FUNCTION_BLOCK PID_SINGLE_UPDATE_SEQUENCE (* One tuning attempt between samples; native validation pending *)
  (* Standard: 61499-2 *)
  (* Version 0.1, 2026-10-24, Guilherme *)
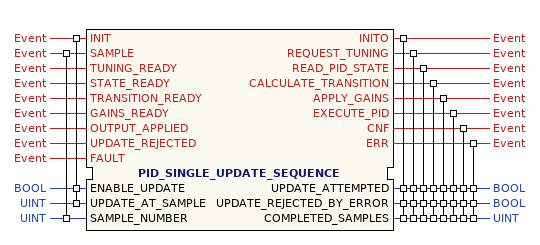
  EVENT_INPUT
    INIT WITH ENABLE_UPDATE, UPDATE_AT_SAMPLE;
    SAMPLE WITH SAMPLE_NUMBER;
    TUNING_READY;
    STATE_READY;
    TRANSITION_READY;
    GAINS_READY;
    OUTPUT_APPLIED;
    UPDATE_REJECTED;
    FAULT;
  END_EVENT
  EVENT_OUTPUT
    INITO WITH UPDATE_ATTEMPTED, UPDATE_REJECTED_BY_ERROR, COMPLETED_SAMPLES;
    REQUEST_TUNING WITH UPDATE_ATTEMPTED, UPDATE_REJECTED_BY_ERROR, COMPLETED_SAMPLES;
    READ_PID_STATE WITH UPDATE_ATTEMPTED, UPDATE_REJECTED_BY_ERROR, COMPLETED_SAMPLES;
    CALCULATE_TRANSITION WITH UPDATE_ATTEMPTED, UPDATE_REJECTED_BY_ERROR, COMPLETED_SAMPLES;
    APPLY_GAINS WITH UPDATE_ATTEMPTED, UPDATE_REJECTED_BY_ERROR, COMPLETED_SAMPLES;
    EXECUTE_PID WITH UPDATE_ATTEMPTED, UPDATE_REJECTED_BY_ERROR, COMPLETED_SAMPLES;
    CNF WITH UPDATE_ATTEMPTED, UPDATE_REJECTED_BY_ERROR, COMPLETED_SAMPLES;
    ERR WITH UPDATE_ATTEMPTED, UPDATE_REJECTED_BY_ERROR, COMPLETED_SAMPLES;
  END_EVENT
  VAR_INPUT
    ENABLE_UPDATE : BOOL;
    UPDATE_AT_SAMPLE : UINT;
    SAMPLE_NUMBER : UINT;
  END_VAR
  VAR_OUTPUT
    UPDATE_ATTEMPTED : BOOL;
    UPDATE_REJECTED_BY_ERROR : BOOL;
    COMPLETED_SAMPLES : UINT;
  END_VAR
  VAR
    RUN_UPDATE_ENABLED : BOOL;
    TARGET_SAMPLE : UINT;
    CURRENT_SAMPLE : UINT;
    INPUT_VALID : BOOL;
    UPDATE_DUE : BOOL;
  END_VAR
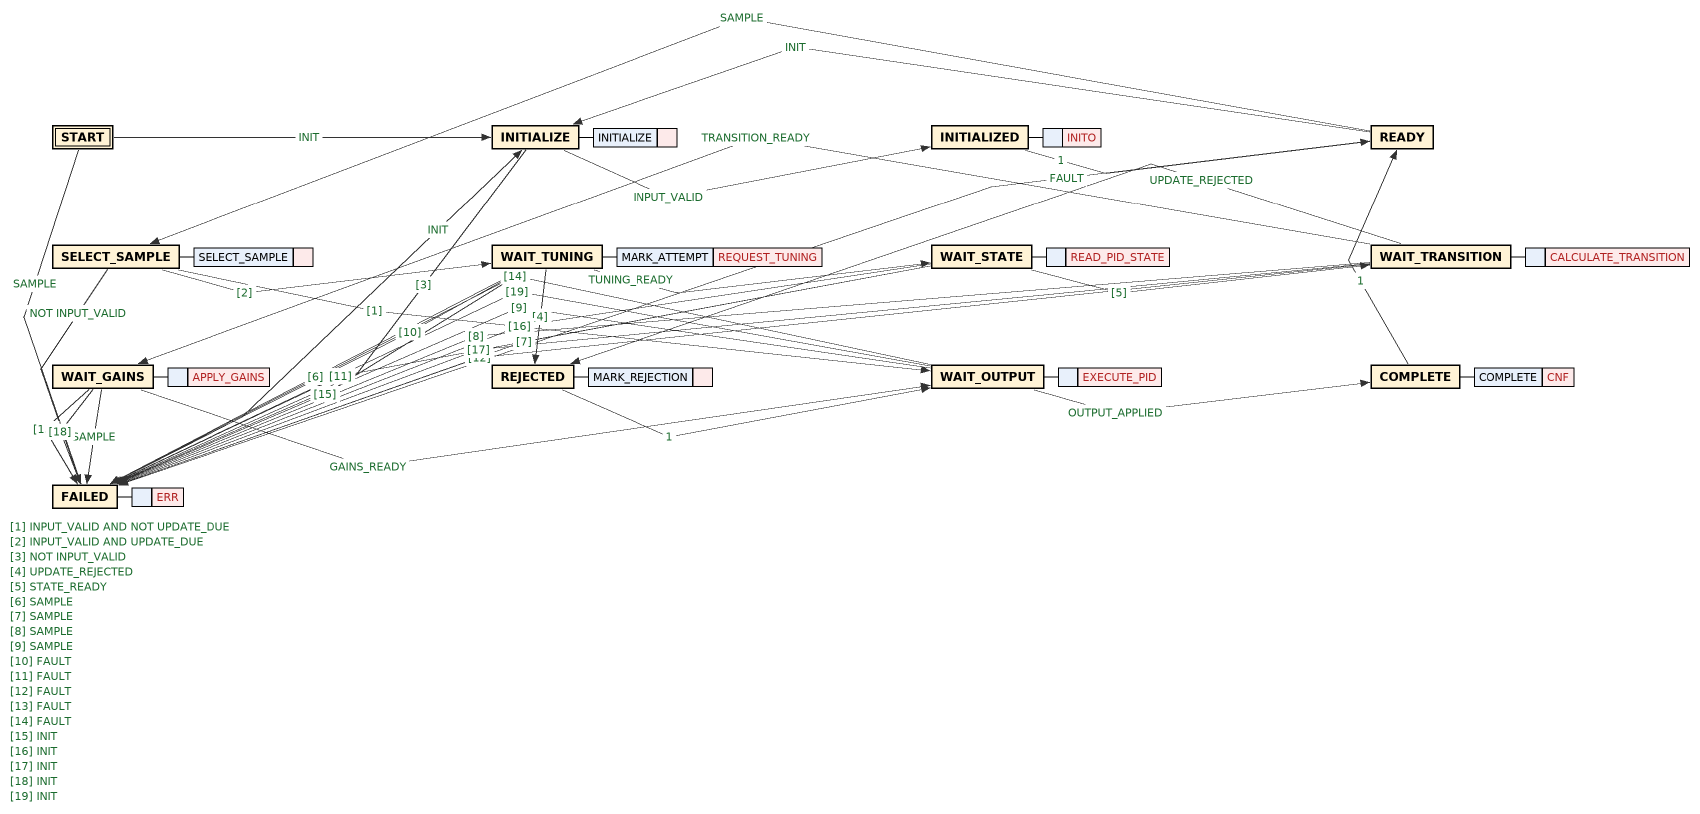
  EC_STATES
    START;
    INITIALIZE : INITIALIZE;
    INITIALIZED : -> INITO;
    READY;
    SELECT_SAMPLE : SELECT_SAMPLE;
    WAIT_TUNING : MARK_ATTEMPT -> REQUEST_TUNING;
    WAIT_STATE : -> READ_PID_STATE;
    WAIT_TRANSITION : -> CALCULATE_TRANSITION;
    WAIT_GAINS : -> APPLY_GAINS;
    REJECTED : MARK_REJECTION;
    WAIT_OUTPUT : -> EXECUTE_PID;
    COMPLETE : COMPLETE -> CNF;
    FAILED : -> ERR;
  END_STATES
  EC_TRANSITIONS
    START TO INITIALIZE := INIT;
    READY TO INITIALIZE := INIT;
    FAILED TO INITIALIZE := INIT;
    START TO FAILED := SAMPLE;
    INITIALIZE TO INITIALIZED := INPUT_VALID;
    INITIALIZE TO FAILED := NOT INPUT_VALID;
    INITIALIZED TO READY := 1;
    READY TO SELECT_SAMPLE := SAMPLE;
    SELECT_SAMPLE TO FAILED := NOT INPUT_VALID;
    SELECT_SAMPLE TO WAIT_TUNING := INPUT_VALID AND UPDATE_DUE;
    SELECT_SAMPLE TO WAIT_OUTPUT := INPUT_VALID AND NOT UPDATE_DUE;
    WAIT_TUNING TO WAIT_STATE := TUNING_READY;
    WAIT_STATE TO WAIT_TRANSITION := STATE_READY;
    WAIT_TRANSITION TO WAIT_GAINS := TRANSITION_READY;
    WAIT_GAINS TO WAIT_OUTPUT := GAINS_READY;
    WAIT_TUNING TO REJECTED := UPDATE_REJECTED;
    WAIT_TRANSITION TO REJECTED := UPDATE_REJECTED;
    REJECTED TO WAIT_OUTPUT := 1;
    WAIT_OUTPUT TO COMPLETE := OUTPUT_APPLIED;
    COMPLETE TO READY := 1;
    WAIT_TUNING TO FAILED := SAMPLE;
    WAIT_TUNING TO FAILED := INIT;
    WAIT_TUNING TO FAILED := FAULT;
    WAIT_STATE TO FAILED := SAMPLE;
    WAIT_STATE TO FAILED := INIT;
    WAIT_STATE TO FAILED := FAULT;
    WAIT_TRANSITION TO FAILED := SAMPLE;
    WAIT_TRANSITION TO FAILED := INIT;
    WAIT_TRANSITION TO FAILED := FAULT;
    WAIT_GAINS TO FAILED := SAMPLE;
    WAIT_GAINS TO FAILED := INIT;
    WAIT_GAINS TO FAILED := FAULT;
    WAIT_OUTPUT TO FAILED := SAMPLE;
    WAIT_OUTPUT TO FAILED := INIT;
    WAIT_OUTPUT TO FAILED := FAULT;
    READY TO FAILED := FAULT;
  END_TRANSITIONS
  ALGORITHM INITIALIZE IN ST:
RUN_UPDATE_ENABLED := ENABLE_UPDATE;
TARGET_SAMPLE := UPDATE_AT_SAMPLE;
CURRENT_SAMPLE := 0;
COMPLETED_SAMPLES := 0;
UPDATE_ATTEMPTED := FALSE;
UPDATE_REJECTED_BY_ERROR := FALSE;
UPDATE_DUE := FALSE;
INPUT_VALID := (NOT RUN_UPDATE_ENABLED) OR (TARGET_SAMPLE > 0);
  END_ALGORITHM
  ALGORITHM SELECT_SAMPLE IN ST:
CURRENT_SAMPLE := SAMPLE_NUMBER;
INPUT_VALID := (CURRENT_SAMPLE > 0) AND (CURRENT_SAMPLE = COMPLETED_SAMPLES + 1);
UPDATE_DUE := RUN_UPDATE_ENABLED AND (NOT UPDATE_ATTEMPTED) AND (CURRENT_SAMPLE = TARGET_SAMPLE);
  END_ALGORITHM
  ALGORITHM MARK_ATTEMPT IN ST:
UPDATE_ATTEMPTED := TRUE;
  END_ALGORITHM
  ALGORITHM MARK_REJECTION IN ST:
UPDATE_REJECTED_BY_ERROR := TRUE;
  END_ALGORITHM
  ALGORITHM COMPLETE IN ST:
COMPLETED_SAMPLES := CURRENT_SAMPLE;
  END_ALGORITHM
END_FUNCTION_BLOCK
